// ST_CylinderParCfg as Modules 0.12 and earlier stored it (v1): the record an
// upgraded station's recipe store still holds, which v2 must refuse (§3.8).
TYPE ST_ProbeCylinderParCfgV1 :
STRUCT
    SchemaVersion : UINT := 1;
    MoveTimeout   : TIME := T#2S;
END_STRUCT
END_TYPE

(* stored: Version 1.1.0.1, ProductVersion 3.1.4024.12
   DUT ST_ProbeCylinderParCfgV1: Id {fe470b9d-beee-408d-9fc5-b5924e6c67f1} *)
